(* Additional processing to handle clocks - in CODESYS, it only starts
    with rising edge and can not be placed inside IF statement *) 
IF(t0_up = TRUE) THEN
    t0_reset := TRUE;
ELSIF(t0_start = TRUE AND t0_up = FALSE) THEN
    t0_up := TRUE;  t0_reset := FALSE;
END_IF
t0(IN:=t0_reset, PT:=T0_VALUE); 
IF(t1_up = TRUE) THEN
    t1_reset := TRUE;
ELSIF(t1_start = TRUE AND t1_up = FALSE) THEN
    t1_up := TRUE;  t1_reset := FALSE;
END_IF
t1(IN:=t1_reset, PT:=T1_VALUE);

END_FUNCTION_BLOCK
